{attribute 'qualified_only'}
{attribute 'strict'}
{attribute 'to_string'}
TYPE E_LogRecordExporterState :
(
	SUCCESS := 0,
	BUSY,
	FAILURE
);
END_TYPE

(* stored: Version 1.1.0.1
   EnumerationTextList E_LogRecordExporterState: Id {dc414b3e-ec7f-4e45-b7f0-3326c54a2985} *)
